(* IEC 61131-3 sources: plcassist-cli/packages/volt-lsp-iec/test-corpus/pro2193/Device/Plc Logic/Application/09 Misc/Library Manager/(unresolved)/iodriver profibus2 interfaces, 7 files *)

(* ---- INTERFACEIDS.gvl ---- *)
VAR_GLOBAL
	ITFID_ICMPIODRVPROFIBUS : DWORD := 16#32;
	ITFID_ICMPIODRVPBSLAVEACTIVATION : DWORD := 16#50;
	ITFID_ICMPIODRVPROFIBUSCONFIG : DWORD := 16#5A;
END_VAR

(* ---- OPERATIONSTATES.gvl ---- *)
VAR_GLOBAL
	PB_NOT_ENABLED : WORD := 0;
	PB_INVALID_PARAMETER : WORD := 1;
	PB_PENDING : WORD := 2;
	PB_DONE : WORD := 3;
	PB_ERROR : WORD := 4;
END_VAR

(* ---- SLAVEACTIVATIONCOMMANDS.gvl ---- *)
VAR_GLOBAL
	PB_SLAVE_ACTIVE : UDINT := 0;
	PB_SLAVE_INACTIVE : UDINT := 1;
END_VAR

(* ---- ICMPIODRVPBSLAVEACTIVATION.itf ---- *)
INTERFACE ICMPIODRVPBSLAVEACTIVATION
END_INTERFACE

METHOD GETSLAVEACTIVATION : UDINT
VAR_IN_OUT
	TSLAVEACTIVATION : PB_SlaveActivation;
END_VAR
END_METHOD

METHOD SETSLAVEACTIVATION : UDINT
VAR_IN_OUT
	TSLAVEACTIVATION : PB_SlaveActivation;
END_VAR
END_METHOD

(* ---- ICMPIODRVPROFIBUS.itf ---- *)
INTERFACE ICMPIODRVPROFIBUS
END_INTERFACE

METHOD CLEARDATA : UDINT
VAR_INPUT
	UDIREMADR : UDINT;
	UDIGROUPSELECT : UDINT;
END_VAR
END_METHOD

METHOD FREEZE : UDINT
VAR_INPUT
	UDIREMADR : UDINT;
	UDIGROUPSELECT : UDINT;
END_VAR
END_METHOD

METHOD SYNC : UDINT
VAR_INPUT
	UDIREMADR : UDINT;
	UDIGROUPSELECT : UDINT;
END_VAR
END_METHOD

METHOD UNSYNC : UDINT
VAR_INPUT
	UDIREMADR : UDINT;
	UDIGROUPSELECT : UDINT;
END_VAR
END_METHOD

METHOD UNFREEZE : UDINT
VAR_INPUT
	UDIREMADR : UDINT;
	UDIGROUPSELECT : UDINT;
END_VAR
END_METHOD

(* ---- ICMPIODRVPROFIBUSCONFIG.itf ---- *)
INTERFACE ICMPIODRVPROFIBUSCONFIG
END_INTERFACE

METHOD GETSLAVECONFIGURATION : UDINT
VAR_IN_OUT
	TGETSLAVECONFIG : PB_SlaveConfigurationData;
END_VAR
END_METHOD

(* ---- IPBSLAVEDIAG.itf ---- *)
INTERFACE IPBSLAVEDIAG
END_INTERFACE

METHOD GETDIAG : DPSlaveDiag
END_METHOD

METHOD GETEXTDIAG : UINT
VAR_INPUT
	PEXTDIAG : POINTER TO BYTE;
	UIMAXLEN : UINT;
END_VAR
END_METHOD
